TYPE (* logiBUS PI Struct Octal *)
  (* Version 1.0, 2026-05-28, franz *)
  PACKAGE logiBUS::io::PI;
  IMPORT logiBUS::io::PI::logiBUS_PI_S;
  logiBUS_PI_S_Octal : STRUCT
    Port1 : logiBUS_PI_S := (Pin := 255);
    Port2 : logiBUS_PI_S := (Pin := 255);
    Port3 : logiBUS_PI_S := (Pin := 255);
    Port4 : logiBUS_PI_S := (Pin := 255);
    Port5 : logiBUS_PI_S := (Pin := 255);
    Port6 : logiBUS_PI_S := (Pin := 255);
    Port7 : logiBUS_PI_S := (Pin := 255);
    Port8 : logiBUS_PI_S := (Pin := 255);
  END_STRUCT;
END_TYPE
